(* CODESYS project settings.library
   DefaultNamespace: KOSTAL.TC3.Core.Settings
   Description: Contains  KOSTAL Framework Global Settinhs
   Author: Frank Dümpelmann
   DocFormat: reStructuredText
   Title: KOSTAL.TC3.Core.Settings
   Version: 2019.0.1.0
   Company: KOSTAL GmbH & Co.KG
   Placeholder: KOSTAL.TC3.Core.Settings

Project tree, tasks and I/O mapping:
  DUT/
    data type T_MaxString
  Project Information/
    function F_GetCompany [ST]
    function F_GetTitle [ST]
    function F_GetVersion [ST]
  Version/
    global variables Global_Version
  global variables CORE_GVL
*)

// DUT/T_MaxString
TYPE T_MaxString : STRING[255]; END_TYPE

// Version/Global_Version
{attribute 'TcGenerated'}
{attribute 'no-analysis'}
{attribute 'linkalways'}
// This function has been automatically generated from the project information.
VAR_GLOBAL CONSTANT
	{attribute 'const_non_replaced'}
	stLibVersion_KOSTAL_TC3_Core_Settings : ST_LibVersion := (iMajor := 2019, iMinor := 0, iBuild := 1, iRevision := 0, nFlags := 0, sVersion := '2019.0.1.0');
END_VAR

// CORE_GVL
{attribute 'qualified_only'}
{attribute 'global_init_slot' := '40010'}
VAR_GLOBAL CONSTANT
	MAX_STRING_LENGHT	:	INT:= 255; // INT:= 255
END_VAR

// Project Information/F_GetCompany
// This function has been automatically generated from the project information.
{attribute 'signature_flag' := '1073741824'}
{attribute 'TcGenerated'}
{attribute 'no-analysis'}
FUNCTION F_GetCompany : WSTRING
VAR_INPUT
	
END_VAR

F_GetCompany := "KOSTAL GmbH & Co.KG";

END_FUNCTION

// Project Information/F_GetTitle
// This function has been automatically generated from the project information.
{attribute 'signature_flag' := '1073741824'}
{attribute 'TcGenerated'}
{attribute 'no-analysis'}
FUNCTION F_GetTitle : WSTRING
VAR_INPUT
	
END_VAR

F_GetTitle := "KOSTAL.TC3.Core.Settings";

END_FUNCTION

// Project Information/F_GetVersion
// This function has been automatically generated from the project information.
{attribute 'signature_flag' := '1073741824'}
{attribute 'TcGenerated'}
{attribute 'no-analysis'}
FUNCTION F_GetVersion : ST_LibVersion
VAR_INPUT
	
END_VAR

F_GetVersion.iMajor := 2019;
F_GetVersion.iMinor := 0;
F_GetVersion.iBuild := 1;
F_GetVersion.iRevision := 0;

END_FUNCTION
